{attribute 'pack_mode' := '1'}
TYPE ST_ScheduleHoliday_V1 :
STRUCT
 Name : STRING(20);
 Priority : UDINT;
 StartDate : UDINT;
 EndDate : UDINT;
END_STRUCT
END_TYPE

(* stored: Version 1.1.0.1, ProductVersion 3.1.4024.15
   DUT ST_ScheduleHoliday_V1: Id {c12ca363-f0a9-4b27-8070-d46bbe3e35fd} *)
